(* IEC 61131-3 sources: codesys-to-s7/tests/corpus/C2S7-ADDR-OVERLAP/pos, 1 file *)

(* ---- input.st ---- *)
VAR_GLOBAL
    wStat AT %MW5 : WORD;
    xBit AT %MX10.0 : BOOL;
END_VAR
